// TIA Portal V21 export
// export: Created 2026-08-21T20:18:56.6880349Z, ExportSetting None, DisplayName Totally Integrated Automation Portal, DisplayVersion V21, DisplayName STEP 7 Professional, DisplayVersion V21, DisplayName STEP 7 Safety, DisplayVersion V21, DisplayName Tech WebApplication, DisplayVersion V21, DisplayName WinCC Basic/Comfort/Advanced, DisplayVersion V21, DisplayName WinCC Professional, DisplayVersion V21, DisplayName WinCC Unified, DisplayVersion V21
TYPE "UDT_Service_StepOrderRawDataMedium"
   STRUCT
      stepOrder : Array[0..199] of "UDT_Service_StepOrder";
      parameterIndex : Array[0..511] of Byte;
   END_STRUCT;
END_TYPE
